// TIA Portal V21 export
VAR_GLOBAL   // PLC tag table "Tags_Filling"
   FillValveOpen AT %Q4.0 : Bool;   // Filling valve open
   FillLevelHigh AT %I4.0 : Bool;   // Filling level high
   FillFlowRaw AT %IW6 : Word;   // Raw value of the filling flow
END_VAR
